Fanuc KAREL source: kt00415.KL

-- PROVISIONAL review KL for V770-1; original PC SHA256 6457374408e21d44fdb1d4ae651aacb02da1e3e077f6500d2f324ce730ff58c1
-- Incomplete behavior may be omitted. Consult companion uncertainty JSON. Do not deploy.
PROGRAM KT00415
%NOLOCKGROUP
VAR
  I2 : INTEGER
  OUT : BOOLEAN
-- UNRESOLVED_DECL H1 type=002017
BEGIN
  -- UNRESOLVED_PC offsets 5-19; opcodes 2E,22,9D,33,B4
  -- UNRESOLVED_PC offsets 24-35; opcodes 2E,23
  -- UNRESOLVED_PC offsets 40-62; opcodes 22,9D,33,B3,21,5B,23
  -- UNRESOLVED_PC offsets 67-71; opcodes 7F
END KT00415
